Staubli VAL3: click_RotHome.pgx

program click_RotHome()
  local bool l_bResult
begin
  if workingMode()!=1
    popUpMsg("非手动模式不支持路径回原！")
    return
  endIf
  //手动机器人路径回原
  l_bResult=userPageConfirm("确认原路径返回Home？")
  if l_bResult
    rs:nCycleCmd=7
    delay(0.2)
    rs:nCycleCmd=0
  endIf

end
